Staubli VAL3: taskManager.pgx

program taskManager()
begin
  //任务守护：某个任务因通信中断/异常退出后，5 秒后自动拉起
  do
    if taskStatus("stateMachine")!=1
      taskResume("stateMachine",1)
      delay(5)
    endIf
    delay(0)
  until false
end
